{attribute 'enable_dynamic_creation'}
FUNCTION_BLOCK FB_SpanId IMPLEMENTS I_OtlpValue
VAR_OUTPUT
	bytes: ARRAY [0..7] OF BYTE;
END_VAR

(*
	Releases this value and clears the caller's pointer to it: call it as p^.delete(pSelf:=p).
	pSelf is cleared before the value is freed, so the caller never keeps a dangling pointer.
	A pointer to any other object is refused and left untouched, and nothing is released.
*)
METHOD delete : BOOL
VAR_IN_OUT
	pSelf: POINTER TO FB_SpanId;
END_VAR
VAR
	_pThis: POINTER TO FB_SpanId;
END_VAR
_pThis := THIS;
IF pSelf <> _pThis THEN
	RETURN;
END_IF

pSelf := 0;
__DELETE(_pThis);
delete := TRUE;
END_METHOD

PROPERTY eType : E_ValueType
GET
eType := E_ValueType.E_SpanId;
END_GET
END_PROPERTY

//FB_Exit must be implemented explicitly. If there is an implementation, then the
//method is called before the controller removes the code of the function block instance
//(implicit call). The return value is not evaluated.
METHOD FB_Exit: BOOL
VAR_INPUT
    bInCopyCode: BOOL;  // TRUE: the exit method is called in order to leave the instance which will be copied afterwards (online change).  
END_VAR
THIS^.free();
END_METHOD

(* deallocates all data owned by the value without deleting the object itself.*)
METHOD free
MEMSET(ADR(THIS^.bytes), 0, SIZEOF(THIS^.bytes));
END_METHOD

END_FUNCTION_BLOCK

(* stored: Version 1.1.0.1
   POU FB_SpanId: Id {5bf3062c-d603-43ca-8490-cc9822c82385}, SpecialFunc None
   Method delete: Id {e7cda35d-3a46-47f9-bedc-fb9f4eebf05c}
   Property eType: Id {386b755d-4227-473a-8d9f-1dcee7cc6d49}
   Get Get: Id {43f7c6c3-7397-4194-ac11-7e0b8b201aec}
   Method FB_Exit: Id {b7cf1790-e849-49d8-a0f6-942cd887bf9e}
   Method free: Id {9d4a26f9-0175-4cf4-a756-1effe28ccc8b} *)
